INTERFACE I_Sample EXTENDS __System.IQueryInterface

METHOD Execute : BOOL
VAR_INPUT
    nMode : INT;
END_VAR
END_METHOD

PROPERTY Busy : BOOL
GET
END_GET
END_PROPERTY

END_INTERFACE

(* stored: Version 1.1.0.1, ProductVersion 3.1.4024.12
   Itf I_Sample: Id {11111111-2222-3333-4444-888888888888}
   Method Execute: Id {bbbbbbbb-0000-0000-0000-000000000001}
   Property Busy: Id {bbbbbbbb-0000-0000-0000-000000000002}
   Get Get: Id {bbbbbbbb-0000-0000-0000-000000000003} *)
